// TIA Portal V21 export
TagTable "T_V6"
  X_V6 :   (PLC tag HMI_IF.SwOn, HMI_Connection_1)
